(* IEC 61131-3 sources: s7-to-codesys/src/GVLs/Converted, 6 files *)

(* ---- DB_Hmi.gvl.st ---- *)
// Назначение: HMI interface
// Автор:      WTP2 (исходный блок S7); перевод в ST — s7conv 0.1.0
// Версия:     0.2 (исходный блок S7)
// Документ:   docs/CONVERSION_REPORT.md, docs/MAPPING.md
// Источник:   samples/scl/DB_Plant.scl, строки 81–109, DATA_BLOCK "DB_Hmi", FAMILY Hmi
// Сгенерировано s7conv: пометки MIGRATION-CHECK и MIGRATION-TODO требуют ручного разбора.
{attribute 'qualified_only'}
VAR_GLOBAL
    cmdWord : WORD;  // Запросы режима (биты, см. FB_ModeSelect); ФБ сбрасывает обработанные биты
    modeRequest : INT := -1;  // Запрос режима числом: -1 — нет запроса
    pump : ARRAY[1..3] OF ST_DB_Hmi_pump;
    alarmAck : BOOL;  // Квитирование аварий
    backwashStart : BOOL;  // Пуск промывки фильтра
    backwashStop : BOOL;  // Прерывание промывки
    resetTotal : BOOL;  // Сброс сменного счётчика объёма
    setpointPressure : REAL := 4.5;  // Уставка давления в коллекторе, бар
    pidManual : BOOL;  // Ручной режим регулятора давления
    pidManualValue : REAL;  // Ручное задание частоты, %
    message : STRING(20);  // Текст для бегущей строки
END_VAR

(* ---- DB_Plant.gvl.st ---- *)
// Назначение: Plant process data
//             Технологические данные станции II подъёма
// Автор:      WTP2 (исходный блок S7); перевод в ST — s7conv 0.1.0
// Версия:     0.3 (исходный блок S7)
// Документ:   docs/CONVERSION_REPORT.md, docs/MAPPING.md
// Источник:   samples/scl/DB_Plant.scl, строки 29–79, DATA_BLOCK "DB_Plant", FAMILY Plant
// Сгенерировано s7conv: пометки MIGRATION-CHECK и MIGRATION-TODO требуют ручного разбора.
// ---- комментарий в начале исходного файла SCL ----
// =============================================================================
// s7-to-codesys — корпус SCL. Написан с нуля, объект вымышленный (ВОС «Северная»).
//
// Файл:   DB_Plant.scl
// Блоки:  глобальные DB "DB_Plant", "DB_Hmi", "DB_Telegram";
//         DB по типу UDT "DB_RecipeActive";
//         экземплярные DB функциональных блоков (18 шт.).
// -----------------------------------------------------------------------------
// Назначение
//   Все блоки данных станции в одном исходнике («Generate source from blocks»
//   для группы DB). Логики нет, кроме начальных значений в секции BEGIN.
//   DB_Plant        — технологические данные; часть переменных сохраняемая
//                     (секция VAR RETAIN): объём за всё время, наработка
//                     фильтров, число промывок.
//   DB_Hmi          — интерфейс с панелью оператора: команды, уставки, текст.
//   DB_Telegram     — неоптимизированный DB (S7_Optimized_Access := 'FALSE')
//                     с фиксированной раскладкой байтов: к нему обращаются
//                     абсолютно (%DB30.DBW0, P#DB30.DBX4.0) и через PEEK/POKE.
//                     Номер DB30 — свойство блока, в исходник TIA не попадает
//                     (см. BlockProperties.csv).
//   DB_RecipeActive — DB, созданный по типу "UDT_DosingRecipe". По тексту его
//                     не отличить от экземплярного DB: нужна таблица символов.
//   Экземплярные DB записаны в двух формах: как выгружает TIA Portal (имя ФБ
//   отдельной строкой после NON_RETAIN) и компактно (DATA_BLOCK "DB" "FB").
// Что проверяет при конвертации
//   DB -> GVL; RETAIN -> RETAIN/PERSISTENT; экземплярный DB -> экземпляр ФБ в GVL;
//   начальные значения из BEGIN; массив UDT; DTL (нет аналога в CODESYS Standard).
// =============================================================================
{attribute 'qualified_only'}
VAR_GLOBAL
    estopOk : BOOL;  // Аварийный стоп не нажат (копия %I0.0)
    tankLevel : REAL := 0.0;  // Уровень в РЧВ, м
    flowSamples : ARRAY[1..8] OF REAL;  // Выборка расхода FT101 раз в секунду, м3/ч
    flowMin : REAL;  // Минимум по выборке, м3/ч
    flowMax : REAL;  // Максимум по выборке, м3/ч
    flowAvg : REAL;  // Среднее по выборке, м3/ч
    flowSampleCount : INT;  // Число достоверных отсчётов в выборке
    clockMem : BOOL;  // Память фронта меркера тактов "Clock_1Hz"
    pressureCfg : UDT_AnalogCfg := (rangeHigh := 16.0);  // Параметры канала PT101 для HMI
    pumpStatus : ARRAY[1..3] OF UDT_DeviceStatus;  // Состояния насосов P101...P103
    plantMode : INT := 1;  // 0 — стоп, 1 — работа, 2 — промывка
    alarmWord : WORD;  // Слово аварий станции (биты см. OB "Main")
    alarmDWord : DWORD;  // Расширенное слово аварий
    heartbeat : BYTE;  // Счётчик жизни для верхнего уровня
    pressureFastRaw : INT;  // Давление PT101, прямое чтение периферии
    lastStart : DT;  // Время последнего пуска станции
    // MIGRATION-TODO: DTL — структура S7 (YEAR, MONTH, ...), в CODESYS нет; заменить на DT или свою структуру (стр.
    //                 53)
    // defaultClock { ExternalAccessible := 'False'; ExternalVisible := 'False'; ExternalWritable := 'False'} : DTL;
    clockLost : BOOL;  // Часы CPU потеряны при запуске
    diagCount : DINT;  // Число диагностических прерываний
    diagLastLaddr : WORD;  // Аппаратный идентификатор последнего модуля с диагностикой
    diagLastChannel : UINT;  // Канал последней диагностики
    diagIoState : WORD;  // IO_State последней диагностики
    operatorName : STRING(20) := 'NOBODY';  // Оператор смены
    shiftData : ST_DB_Plant_shiftData;
END_VAR
VAR_GLOBAL RETAIN
    totalVolume : LREAL;  // Объём за всё время, м3 (копия из DB_FQ101)
    filterRuntime : ARRAY[1..4] OF TIME;  // Наработка фильтров с последней промывки
    backwashCount : DINT;  // Число промывок
END_VAR

(* ---- DB_Telegram.gvl.st ---- *)
// Назначение: Legacy telegram buffer
//             Буфер телеграммы удалённой станции (раскладка байтов фиксирована: DBW0 заголовок, DBW2 номер,
//             DBB4...19 данные)
// Автор:      WTP1 (исходный блок S7); перевод в ST — s7conv 0.1.0
// Версия:     1.1 (исходный блок S7)
// Документ:   docs/CONVERSION_REPORT.md, docs/MAPPING.md
// Источник:   samples/scl/DB_Plant.scl, строки 111–131, DATA_BLOCK "DB_Telegram", FAMILY Comm
// Сгенерировано s7conv: пометки MIGRATION-CHECK и MIGRATION-TODO требуют ручного разбора.
// MIGRATION-CHECK: стандартный (неоптимизированный) доступ S7: абсолютная адресация и порядок байтов не переносятся
//                  (стр. 111)
{attribute 'qualified_only'}
VAR_GLOBAL
    header : WORD;  // DBW0: слово состояния станции
    seqNo : WORD;  // DBW2: номер телеграммы
    payload : ARRAY[0..15] OF BYTE;  // DBB4...DBB19: данные
    crc : WORD;  // DBW20
    reserve : ARRAY[0..12] OF BYTE;  // DBB22...DBB34
    heartbeat : BYTE;  // DBB35: счётчик жизни (пишет POKE в FB_EventLogger)
END_VAR

(* ---- GVL_InstanceDBs.gvl.st ---- *)
// Назначение: экземпляры функциональных блоков и типизированные DB S7 (экземплярные DB → переменные GVL)
// Автор:      s7conv 0.1.0 (сгенерировано)
// Версия:     не указана
// Документ:   docs/MAPPING.md, раздел «DB»
{attribute 'qualified_only'}
VAR_GLOBAL
    DB_AlarmPT101 : FB_AlarmDelay; // samples/scl/DB_Plant.scl:236
    DB_Backwash : FB_Sequencer := (drainTimeout := T#90S); // samples/scl/DB_Plant.scl:200
    DB_Dosing : FB_BatchCounter := (pulsesPerDose := 50); // samples/scl/DB_Plant.scl:257
    DB_FQ101 : FB_Totalizer := (lowFlowCutoff := 2.0); // samples/scl/DB_Plant.scl:190
    DB_FT101 : FB_AnalogIn := (rangeHigh := 1200.0,
                               limitHH := 1150.0,
                               limitH := 1100.0,
                               limitL := 0.0,
                               limitLL := -1.0,
                               hysteresis := 10.0); // samples/scl/DB_Plant.scl:226
    DB_Logger : FB_EventLogger; // samples/scl/DB_Plant.scl:262
    DB_LS201 : FB_Debounce; // samples/scl/DB_Plant.scl:248
    DB_LT101 : FB_AnalogIn := (rangeHigh := 5.0,
                               limitHH := 4.8,
                               limitH := 4.5,
                               limitL := 1.0,
                               limitLL := 0.5,
                               hysteresis := 0.05); // samples/scl/DB_Plant.scl:216
    DB_Mode : FB_ModeSelect; // samples/scl/DB_Plant.scl:240
    DB_P101 : FB_Motor := (feedbackTime := T#5S); // samples/scl/DB_Plant.scl:146
    DB_P102 : FB_Motor := (feedbackTime := T#5S); // samples/scl/DB_Plant.scl:157
    DB_P103 : FB_Motor; // samples/scl/DB_Plant.scl:168
    DB_PIC101 : FB_PIController := (kp := 2.0, ti := T#20S); // samples/scl/DB_Plant.scl:178
    DB_PT101 : FB_AnalogIn := (rangeHigh := 16.0); // samples/scl/DB_Plant.scl:211
    DB_PumpAlt : FB_PumpAlternation; // samples/scl/DB_Plant.scl:244
    DB_RampSP : FB_Ramp; // samples/scl/DB_Plant.scl:270
    DB_RecipeActive : UDT_DosingRecipe := (name := 'SUMMER',
                                           doseStep := [0.8, 1.2, 1.5, 2.0]); // samples/scl/DB_Plant.scl:133
    DB_XV201 : FB_Valve := (travelTime := T#45S); // samples/scl/DB_Plant.scl:252
END_VAR
VAR_GLOBAL RETAIN
    // MIGRATION-CHECK: стандартный (неоптимизированный) экземплярный или типизированный DB без NON_RETAIN: в S7 он
    //                  реманентный целиком — объявлен в VAR_GLOBAL RETAIN GVL_InstanceDBs (стр. 266)
    DB_LegacyTlg : FB_LegacyTelegram; // samples/scl/DB_Plant.scl:266
END_VAR

(* ---- GVL_IO.gvl.st ---- *)
// Назначение: символьный слой входов/выходов S7: прямые адреса и теги с адресом → переменные с AT
// Автор:      s7conv 0.1.0 (сгенерировано)
// Версия:     не указана
// Документ:   docs/MAPPING.md, раздел «Адреса»
// Адресная модель: S7 нумерует байты (%IW64 — байты 64–65, big-endian), CODESYS — слова
// (%IW32 — байты 64–65, little-endian). Адреса ниже — заготовка: на ПЛК210 каналы модулей
// привязываются в дереве устройств (I/O mapping) — сверить с конфигурацией.
{attribute 'qualified_only'}
VAR_GLOBAL
    EStop_Ok AT %IX0.0 : BOOL; // S7 %I0.0; Аварийный стоп не нажат (НЗ цепь)
    P101_Fbk AT %IX0.1 : BOOL; // S7 %I0.1; P101 обратная связь контактора
    P101_ThermalOk AT %IX0.2 : BOOL; // S7 %I0.2; P101 тепловое реле в норме
    P102_Fbk AT %IX0.3 : BOOL; // S7 %I0.3; P102 обратная связь контактора
    P102_ThermalOk AT %IX0.4 : BOOL; // S7 %I0.4; P102 тепловое реле в норме
    LS201_Drained AT %IX0.5 : BOOL; // S7 %I0.5; Поплавок: фильтр опорожнён
    LS202_Full AT %IX0.6 : BOOL; // S7 %I0.6; Поплавок: фильтр заполнен
    P103_Fbk AT %IX0.7 : BOOL; // S7 %I0.7; P103 обратная связь контактора
    Sw_Local AT %IX1.0 : BOOL; // S7 %I1.0; Ключ «Местное» на шкафу
    Btn_Ack AT %IX1.1 : BOOL; // S7 %I1.1; Кнопка «Квитирование» на шкафу
    P103_ThermalOk AT %IX1.2 : BOOL; // S7 %I1.2; P103 тепловое реле в норме
    XV201_Opened AT %IX2.0 : BOOL; // S7 %I2.0; XV201 концевик «открыто»
    XV201_Closed AT %IX2.1 : BOOL; // S7 %I2.1; XV201 концевик «закрыто»
    FQ201_Pulse AT %IX3.0 : BOOL; // S7 %I3.0; Импульсы расходомера реагента (геркон НЗ)
    PT101_Raw AT %IW32 : INT; // S7 %IW64; PT101 давление в коллекторе 4-20 мА (0...16 бар)
    LT101_Raw AT %IW33 : INT; // S7 %IW66; LT101 уровень в РЧВ 4-20 мА (0...5 м)
    FT101_Raw AT %IW34 : INT; // S7 %IW68; FT101 расход в сеть 4-20 мА (0...1200 м3/ч)
    PT101_Fast AT %IW136 : INT; // S7 %IW272; Канал быстрого опроса давления (читается как %IW272:P)
    P101_Run AT %QX0.0 : BOOL; // S7 %Q0.0; P101 контактор
    P102_Run AT %QX0.1 : BOOL; // S7 %Q0.1; P102 контактор
    P103_Run AT %QX0.2 : BOOL; // S7 %Q0.2; P103 контактор
    XV_Drain AT %QX0.4 : BOOL; // S7 %Q0.4; Задвижка сброса промывной воды
    Q_AirBlower AT %QX0.5 : BOOL; // S7 %Q0.5; Воздуходувка промывки
    Q_WashPump AT %QX0.6 : BOOL; // S7 %Q0.6; Промывной насос
    XV201_Open AT %QX1.0 : BOOL; // S7 %Q1.0; XV201 пускатель «открыть»
    XV201_Close AT %QX1.1 : BOOL; // S7 %Q1.1; XV201 пускатель «закрыть»
    Lamp_Alarm AT %QX2.0 : BOOL; // S7 %Q2.0; Лампа «Авария» на шкафу
    VFD_SpeedRef AT %QW40 : INT; // S7 %QW80; Задание частоты ПЧ ведущего насоса (0...27648)
END_VAR

(* ---- GVL_Markers.gvl.st ---- *)
// Назначение: символьный слой меркеров (%M) S7: прямые адреса и теги с адресом → переменные с AT
// Автор:      s7conv 0.1.0 (сгенерировано)
// Версия:     не указана
// Документ:   docs/MAPPING.md, раздел «Адреса»
// Адресная модель: S7 нумерует байты (%IW64 — байты 64–65, big-endian), CODESYS — слова
// (%IW32 — байты 64–65, little-endian). Адреса ниже — заготовка: на ПЛК210 каналы модулей
// привязываются в дереве устройств (I/O mapping) — сверить с конфигурацией.
{attribute 'qualified_only'}
VAR_GLOBAL
    Clock_1Hz AT %MX0.5 : BOOL; // S7 %M0.5; Меркер тактов 1 Гц (байт тактовых меркеров MB0)
    HMI_StatusPT101 AT %MW5 : WORD; // S7 %MW10; Слово состояния PT101 для старой панели
    HMI_P101Running AT %MX12.0 : BOOL; // S7 %M12.0; P101 в работе для старой панели
    HMI_DosingPacked AT %MD5 : DWORD; // S7 %MD20; Счётчики дозирования одним словом
    Tlg_Source AT %MB100 : BYTE; // S7 %MB100; Начало области данных телеграммы (P#M100.0 BYTE 16)
END_VAR
